// TIA Portal V21 export
ScreenTemplate "Tpl"  NonexNone
  ScreenLayer 
    TextField "frm_1" at 0,0 size 1024x79
    TextField "txt_1" at 9,5 size 144x18  Text="LUČKA DIZALICA"
    TextField "txt_2" at 9,23 size 144x12  Text="PLC Challenge 2026 - EESTEC"
    Rectangle "lmp_1" at 155,7 size 7x7
      RangeAppearanceAnimation "RangeAppearanceAnimation"
        tag Heartbeat
        0..0: back #aaaaaa, fore #000000
        1..1: back #28a03c, fore #000000
    Button "btn_1" at 171,5 size 85x31  TextOff="UKLJ. / ISKLJ.", TextOn="UKLJ. / ISKLJ."
      on Press: InvertBit(Tag := SwOn)
    Rectangle "lmp_2" at 261,6 size 12x12
      RangeAppearanceAnimation "RangeAppearanceAnimation"
        tag LampReady
        0..0: back #aaaaaa, fore #000000
        1..1: back #28a03c, fore #000000
    TextField "txt_3" at 275,6 size 59x12  Text="SPREMAN"
    Rectangle "lmp_3" at 261,23 size 12x12
      RangeAppearanceAnimation "RangeAppearanceAnimation"
        tag LampOff
        0..0: back #aaaaaa, fore #000000
        1..1: back #28a03c, fore #000000
    TextField "txt_4" at 275,23 size 59x12  Text="ISKLJUČEN"
    Button "btn_2" at 341,5 size 96x31  TextOff="POČETNO STANJE", TextOn="POČETNO STANJE"
      on Press: SetBit(Tag := BtnInit)
    Button "btn_3" at 448,5 size 85x31  TextOff="AUTOMATSKAMANIPULACIJA", TextOn="AUTOMATSKAMANIPULACIJA"
      on Press: SetBit(Tag := BtnAuto)
    Rectangle "lmp_4" at 448,37 size 85x4
      RangeAppearanceAnimation "RangeAppearanceAnimation"
        tag LampAuto
        0..0: back #aaaaaa, fore #000000
        1..1: back #28a03c, fore #000000
    Button "btn_4" at 536,5 size 96x31  TextOff="POLUAUTOMATSKAMANIPULACIJA", TextOn="POLUAUTOMATSKAMANIPULACIJA"
      on Press: SetBit(Tag := BtnSemi)
    Rectangle "lmp_5" at 536,37 size 96x4
      RangeAppearanceAnimation "RangeAppearanceAnimation"
        tag LampSemi
        0..0: back #aaaaaa, fore #000000
        1..1: back #28a03c, fore #000000
    Button "btn_5" at 636,5 size 75x31  TextOff="RUČNOUPRAVLJANJE", TextOn="RUČNOUPRAVLJANJE"
      on Press: SetBit(Tag := BtnManual)
    Rectangle "lmp_6" at 636,37 size 75x4
      RangeAppearanceAnimation "RangeAppearanceAnimation"
        tag LampManual
        0..0: back #aaaaaa, fore #000000
        1..1: back #28a03c, fore #000000
    Button "btn_6" at 721,5 size 64x31  TextOff="START", TextOn="START"
      on Press: SetBit(Tag := BtnStart)
    Rectangle "lmp_7" at 721,37 size 64x4
      RangeAppearanceAnimation "RangeAppearanceAnimation"
        tag LampRunning
        0..0: back #aaaaaa, fore #000000
        1..1: back #28a03c, fore #000000
    Button "btn_7" at 788,5 size 64x31  TextOff="STOP", TextOn="STOP"
      on Press: SetBit(Tag := BtnStop)
    Button "btn_8" at 855,5 size 64x31  TextOff="POTVRDA", TextOn="POTVRDA"
      on Press: SetBit(Tag := BtnAck)
    Button "btn_9" at 923,5 size 94x31  TextOff="SLJEDEĆI KORAK", TextOn="SLJEDEĆI KORAK"
      on Press: SetBit(Tag := BtnStep)
    Rectangle "lmp_8" at 923,37 size 94x4
      RangeAppearanceAnimation "RangeAppearanceAnimation"
        tag StepWaiting
        0..0: back #aaaaaa, fore #000000
        1..1: back #28a03c, fore #000000
    TextField "txt_5" at 9,49 size 43x18  Text="STANJE"
    SymbolicIOField "sym_1" at 51,49 size 107x18  Mode=Output, TextList=TL_State
      ProcessValue := State
    SymbolicIOField "sym_2" at 161,49 size 95x18  Mode=Output, TextList=TL_Mode
      ProcessValue := Mode
    TextField "txt_6" at 261,49 size 19x18  Text="M"
    IOField "io_1" at 281,49 size 48x18  DataFormat=Decimal, FormatPattern=99999, Mode=Output
      ProcessValue := M
    TextField "txt_7" at 332,49 size 27x18  Text="T [s]"
    IOField "io_2" at 358,49 size 59x18  DataFormat=Decimal, FormatPattern=999999.9, Mode=Output
      ProcessValue := T
    TextField "txt_8" at 421,49 size 14x18  Text="J"
    IOField "io_3" at 435,49 size 48x18  DataFormat=Decimal, FormatPattern=9.9999, Mode=Output
      ProcessValue := J
    TextField "txt_9" at 487,49 size 60x18  Text="Predviđeno"
    IOField "io_4" at 547,49 size 43x18  DataFormat=Decimal, FormatPattern=99999, Mode=Output
      ProcessValue := PredM
    IOField "io_5" at 592,49 size 55x18  DataFormat=Decimal, FormatPattern=999999.9, Mode=Output
      ProcessValue := PredT
    IOField "io_6" at 650,49 size 45x18  DataFormat=Decimal, FormatPattern=9.9999, Mode=Output
      ProcessValue := PredJ
    TextField "txt_10" at 700,49 size 29x18  Text="Trans."
    IOField "io_7" at 728,49 size 28x18  DataFormat=Decimal, FormatPattern=999, Mode=Output
      ProcessValue := TrDone
    TextField "txt_11" at 756,49 size 6x18  Text="/"
    IOField "io_8" at 763,49 size 28x18  DataFormat=Decimal, FormatPattern=999, Mode=Output
      ProcessValue := TrTotal
    Rectangle "lmp_9" at 797,52 size 12x12
      RangeAppearanceAnimation "RangeAppearanceAnimation"
        tag LampAlarm
        0..0: back #aaaaaa, fore #000000
        1..1: back #dc0000, fore #000000, flashing
    SymbolicIOField "sym_3" at 811,49 size 206x18  Mode=Output, TextList=TL_Alarm
      ProcessValue := AlarmHist_00
    TextField "frm_2" at 0,546 size 1024x30
    Button "nav_1" at 9,549 size 107x23  TextOff="GLAVNI PRIKAZ", TextOn="GLAVNI PRIKAZ"
      on Press: ActivateScreen(Screen name := Screen_1, Object number := 0)
    Button "nav_2" at 121,549 size 107x23  TextOff="RUČNO UPRAVLJANJE", TextOn="RUČNO UPRAVLJANJE"
      on Press: ActivateScreen(Screen name := Manual, Object number := 0)
    Button "nav_3" at 233,549 size 107x23  TextOff="LISTE I POSTAVKE", TextOn="LISTE I POSTAVKE"
      on Press: ActivateScreen(Screen name := Lists, Object number := 0)
    Button "nav_4" at 345,549 size 107x23  TextOff="ALARMI", TextOn="ALARMI"
      on Press: ActivateScreen(Screen name := Alarms, Object number := 0)
    Button "nav_5" at 457,549 size 107x23  TextOff="POVIJEST ALARMA", TextOn="POVIJEST ALARMA"
      on Press: ActivateScreen(Screen name := AlarmLog, Object number := 0)
    Button "nav_6" at 568,549 size 117x23  TextOff="REZULTAT / OPTIMIZACIJA", TextOn="REZULTAT / OPTIMIZACIJA"
      on Press: ActivateScreen(Screen name := Score, Object number := 0)
    TextField "txt_12" at 693,551 size 59x18  Text="OB30 takt"
    IOField "io_9" at 752,551 size 59x18  DataFormat=Decimal, FormatPattern=9999999, Mode=Output
      ProcessValue := OB30Ticks
    DateTimeField "dtm_1" at 832,550 size 185x21  Mode=Output
